Universal Robots URScript: SubProg.script

def SubProg():
  # Default parameters:
  global speed_ms = 0.3
  global speed_rads = 0.75
  global accel_mss = 3
  global accel_radss = 1.2
  global blend_radius_m = 0.001

  # Add subprograms here
  # Start of main program
  # Program generated by RoboDK v5.9.4 for UR10 on 26/10/2026 01:01:20
  # Using nominal kinematics.
  # set_reference(p[0.036764, 0.400000, 0.728939, 0.000000, 0.000000, 30.000000])
  set_tcp(p[0.000000, 0.000000, 0.120000, 0.000000, 15.000000, 0.000000])
  movel([-4.065387, -1.176966, 4.792364, -2.498712, 1.044735, -2.370328],accel_mss,speed_ms,0,blend_radius_m)
  # Inside sub
  # End of main program
end

SubProg()
